(* IEC 61131-3 sources: RootPLC/examples/traffic-light/tests, 1 file *)

(* ---- traffic_light_test.st ---- *)
TEST disabled_shows_red_only
VAR
    uut : PRG_TrafficLight;
END_VAR
uut(enable := FALSE);
ASSERT_TRUE(uut.red);
ASSERT_FALSE(uut.yellow OR uut.green);
END_TEST
